// TIA Portal V21 export
DATA_BLOCK "DB_Process"   // DB20
TITLE = Технологические данные (стандартный доступ)
{ S7_Optimized_Access := 'FALSE' }
AUTHOR : WTP2
FAMILY : Plant
VERSION : 0.1
// Неоптимизированный DB: STL S7-300 адресует члены по смещению (Offset)
// stored: AutoNumber false
   VAR
      xPumpRun : Bool;   // Насос в работе
      iLevel_cm : Int;   // Уровень, см
      rFlow_m3h : Real;   // Расход, м3/ч
      wStatus : Word;   // Слово состояния
      stValve : "UDT_Valve";   // Задвижка напорная
   END_VAR
   VAR RETAIN
      iBatch : Int := 1;   // Номер партии
   END_VAR
BEGIN
END_DATA_BLOCK
